Staubli VAL3: logMoveMsgC.pgx

program logMoveMsgC(pointRx x_pPoint1, pointRx x_pPoint2, tool x_tTool, mdesc x_mSpeed, num x_nMoveId)
  local string l_sCode
  local bool l_bResult[2]
  local jointRx l_jRef
  local jointRx l_jResult[2]
begin
  //
  if nRecIndex<200
    // c
    if nRecIndex>=1
      l_jRef=jPointRec[nRecIndex-1,1]
    else
      l_jRef=herej()
    endIf
    l_bResult[0]=pointToJoint(x_tTool,l_jRef,x_pPoint1,l_jResult[0])
    l_bResult[1]=pointToJoint(x_tTool,l_jResult[0],x_pPoint2,l_jResult[1])
    //
    if l_bResult[0]==true and l_bResult[1]==true
      setMutex(bPushToStack)
      jPointRec[nRecIndex,0]=l_jResult[0]
      jPointRec[nRecIndex,1]=l_jResult[1]
      trToolRec[nRecIndex]=x_tTool.trsf
      mSpeedRec[nRecIndex]=x_mSpeed
      nMoveIdRec[nRecIndex]=x_nMoveId
      nMoveTypeRec[nRecIndex]=3
      //logMsg("record moveC."+toString("",nMoveIdRec[nRecIndex]))
      nRecIndex=nRecIndex+1
      bPushToStack=false
    else
      // 无关节解
    endIf
  else
    //popUpMsg("记录点数超过容量.")
  endIf

end
